Staubli VAL3: saveTRAJ.pjx

--- saveTRAJ.pjx ---
Parameters version=s8.10.3Cs9_BS2093 stackSize=5000 millimeterUnit=true
Program file=start.pgx
Program file=stop.pgx
Data file=saveTRAJ.dtx
Type name=trajItem path=Disk://source/template/trajItem/trajItem.pjx

--- saveTRAJ.dtx ---
public trajItem tTrajItem{}
  [Key1]
    pointItem pPointItem
      [0]
        paraItem pParaItem
          [0]
            mdesc mMdesc
            num nMoveType
            num nActionIndex[2]
            num nPercentage[2]
        pointRx pPointRx
        jointRx jJointRx
    num nFrameIndex
    num nToolIndex
    string sID
    num nMoveID

--- start.pgx ---
program start()
begin
end

--- stop.pgx ---
program stop()
begin
end
